(* IEC 61131-3 sources: Test-Git_ESME26/TestProgettoESME_26.fbsproj/PacDriveLib Migration/Motion/MultiCam/PDL_FB_MultiCam.fb.st^/GetPosition, 2 files *)

(* ---- GetCamPositionOfMaster.meth.st ---- *)
METHOD PRIVATE GetCamPositionOfMaster : BOOL
VAR_INPUT
END_VAR

VAR
	etMoinResult				: MOIN.ET_Result;
END_VAR

GetCamPositionOfMaster := TRUE;

etMoinResult :=  MOIN.FC_GetMasterPositionFromGivenSlavePositionForMultiCam(
							i_lrSlavePosition		:= i_ifDrive.lrPosition,
							i_lrMasterScaling		:= 1,
							i_lrSlaveScaling		:= 1,
							i_stCamTableID			:= stActiveMultiCamData,
							i_lrStartPosition		:= iq_stExt.lrXStart,
							i_lrAccuracy			:= iq_stExt.lrAccuracy,
							i_lrIncrementalStepSize	:= iq_stExt.lrXIncr,
							q_lrMasterPosition		=> q_lrPositionX );

IF etMoinResult <> MOIN.ET_Result.Ok THEN

	SetDiagOutput(	i_etDiag	:= GD.ET_Diag.UnexpectedProgramBehavior,
					i_etDiagExt := PDL_ET_DiagExt.UnexpectedFeedback,
					i_sMsg		:= CONCAT('FC_GetMasterPositionFromGivenSlavePositionForMultiCam: ', TO_STRING(etMoinResult)));
	etState := ET_MulticamState.idle_error;
	GetCamPositionOfMaster := FALSE;
	RETURN;
END_IF

(* ---- GetCamPositionOfSlave.meth.st ---- *)
METHOD PRIVATE GetCamPositionOfSlave : BOOL
VAR_INPUT
	i_xCheckModulo			: BOOL;
END_VAR

VAR_OUTPUT
	q_lrSlavePosition		: LREAL;
END_VAR

VAR
	etMoinResult				: MOIN.ET_Result;
	etSetPosResult				: PLCO.ET_Result;
END_VAR

GetCamPositionOfSlave := TRUE;

IF i_xCheckModulo THEN
	IF   q_lrPositionX > stActiveMultiCamData.astCamPoint[0].lrX + lrXPeriode
	  OR q_lrPositionX < stActiveMultiCamData.astCamPoint[0].lrX
	THEN
		//adjust logic encoder position if position is not within period...
		lrModCount := TRUNC_INT((q_lrPositionX - stActiveMultiCamData.astCamPoint[0].lrX) / lrXPeriode);
		IF q_lrPositionX < stActiveMultiCamData.astCamPoint[0].lrX THEN
			lrModCount := lrModCount - 1;
		END_IF
		q_lrPositionX := q_lrPositionX - lrModCount * lrXPeriode;

		fbSetPos( Execute		:= FALSE );
		fbSetPos(	Axis		:= iq_lencMaster,
					Execute		:= TRUE,
					Position	:= - lrModCount * lrXPeriode,
					Relative	:= TRUE,
					ErrorId		=> etSetPosResult );

		IF etSetPosResult <> PLCO.ET_Result.Ok THEN
			SetDiagOutput(	i_etDiag	:= GD.ET_Diag.UnexpectedProgramBehavior,
							i_etDiagExt := PDL_ET_DiagExt.UnexpectedFeedback,
							i_sMsg		:= CONCAT('MC_SetPosition: ', TO_STRING(etSetPosResult)));

			GetCamPositionOfSlave := FALSE;
			etState := ET_MulticamState.idle_error;
			RETURN;
		END_IF

	END_IF
END_IF

//... then get slave cam position
etMoinResult := MOIN.FC_EvaluateMultiCam( 	i_stMultiCam 		:= stActiveMultiCamData,
											i_lrMasterPosition	:= iq_lencMaster.lrPosition,
											q_lrCamPosition		=> q_lrSlavePosition
											);

IF etMoinResult <> MOIN.ET_Result.Ok THEN

	SetDiagOutput(	i_etDiag	:= GD.ET_Diag.UnexpectedProgramBehavior,
					i_etDiagExt	:= PDL_ET_DiagExt.UnexpectedFeedback,
					i_sMsg		:= CONCAT('MOIN.FC_EvaluateMultiCam: ', TO_STRING(etMoinResult)));

	GetCamPositionOfSlave := FALSE;
	etState := ET_MulticamState.idle_error;
	RETURN;
END_IF
